Fanuc KAREL source: ka00120.KL

-- PROVISIONAL review KL for V940-1; original PC SHA256 eb8929a2d270ddbb3253aeaceb2edfee8f53c03c224a2b58aa9cf99e97060c20
-- Incomplete behavior may be omitted. Consult companion uncertainty JSON. Do not deploy.
PROGRAM KA00120
%NOLOCKGROUP
-- UNRESOLVED_DECL SRC type=00001c
-- UNRESOLVED_DECL DST type=002017
BEGIN
  -- V9_ZERO_TABLE_METADATA_HINT layout=0001; no indexed target words; source/name/runtime held
  -- UNRESOLVED_PC offsets 5-15; opcodes 9D,22,A5
  -- UNRESOLVED_PC offsets 20-35; opcodes 21,22,9D,33,B4
  -- UNRESOLVED_PC offsets 40-44; opcodes 7F
END KA00120
